Fanuc KAREL source: kd00020.KL

-- PROVISIONAL review KL for V1013-1; original PC SHA256 2657d865443d5ea117dbf525fd2a7d4723f6b1cbeddc32b80ff6da2b1feed0d4
-- Incomplete behavior may be omitted. Consult companion uncertainty JSON. Do not deploy.
PROGRAM KD00020
%NOLOCKGROUP
VAR
  I : INTEGER
  J : INTEGER
  B : BOOLEAN
  R : REAL
  S : STRING[80]
BEGIN
  -- UNRESOLVED_PC offsets 5-10; opcodes 7A
  -- UNRESOLVED_PC offsets 15-22; opcodes 9D,23
  -- UNRESOLVED_PC offsets 27-31; opcodes 7F
END KD00020
